FUNCTION_BLOCK manual (* Basic Function Block Type *)
  (* Standard: 61499-2 *)
  (* Version 0.0, 10/21/2026, lizar, Schneider Electric, Template *)
  PACKAGE Main;
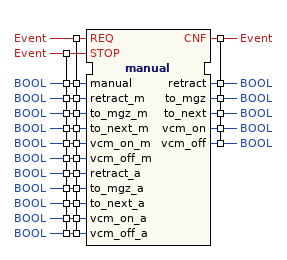
  EVENT_INPUT
    REQ WITH manual, retract_m, to_mgz_m, to_next_m, vcm_on_m, vcm_off_m, retract_a, to_mgz_a, to_next_a, vcm_on_a, vcm_off_a; (* Initialization Request *)
    STOP WITH manual, retract_m, to_mgz_m, to_next_m, vcm_on_m, vcm_off_m, retract_a, to_mgz_a, to_next_a, vcm_on_a, vcm_off_a;
  END_EVENT
  EVENT_OUTPUT
    CNF WITH retract, to_mgz, to_next, vcm_on, vcm_off; (* Execution Confirmation *)
  END_EVENT
  VAR_INPUT
    manual : BOOL;
    retract_m : BOOL;
    to_mgz_m : BOOL;
    to_next_m : BOOL;
    vcm_on_m : BOOL;
    vcm_off_m : BOOL;
    retract_a : BOOL;
    to_mgz_a : BOOL;
    to_next_a : BOOL;
    vcm_on_a : BOOL;
    vcm_off_a : BOOL;
  END_VAR
  VAR_OUTPUT
    retract : BOOL; (* Output event qualifier *)
    to_mgz : BOOL;
    to_next : BOOL;
    vcm_on : BOOL;
    vcm_off : BOOL;
  END_VAR
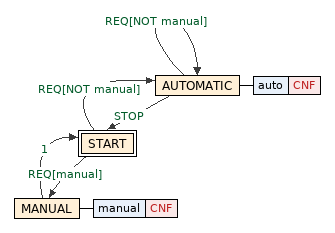
  EC_STATES
    START; (* Initial State *)
    AUTOMATIC : auto -> CNF; (* Initialization *)
    MANUAL : manual -> CNF; (* Normal execution *)
  END_STATES
  EC_TRANSITIONS
    START TO AUTOMATIC := REQ[NOT manual];
    AUTOMATIC TO START := STOP;
    START TO MANUAL := REQ[manual];
    MANUAL TO START := 1;
    AUTOMATIC TO AUTOMATIC := REQ[NOT manual];
  END_TRANSITIONS
  ALGORITHM manual IN ST: (* Initialization algorithm *)
;
retract:=retract_m;
to_mgz:=to_mgz_m;
to_next:=to_next_m;
vcm_on:=vcm_on_m;
vcm_off:=vcm_off_m;
  END_ALGORITHM
  ALGORITHM auto IN ST:
;
retract:=retract_a;
to_mgz:=to_mgz_a;
to_next:=to_next_a;
vcm_on:=vcm_on_a;
vcm_off:=vcm_off_a;
  END_ALGORITHM
END_FUNCTION_BLOCK
